// TIA Portal V21 export
// export: Created 2026-11-11T00:48:17.7043043Z, ExportSetting WithDefaults, DisplayName Totally Integrated Automation Portal, DisplayVersion V21 Update 3, DisplayName STEP 7 Professional, DisplayVersion V21 Update 3, DisplayName STEP 7 Safety, DisplayVersion V21, DisplayName Tech WebApplication, DisplayVersion V21, DisplayName WinCC Basic/Comfort/Advanced, DisplayVersion V21 Update 3, DisplayName WinCC Unified, DisplayVersion V21 Update 3
FUNCTION_BLOCK "FB_Scl_sl053"   // FB31, SCL
{ S7_Optimized_Access := 'TRUE' }
VERSION : 0.1
// stored: AutoNumber true, IsIECCheckEnabled false, IsRetainMemResEnabled false, MemoryReserve 100, SetENOAutomatically false, UDAEnableTagReadback false
   VAR_INPUT
      v_req : Bool;
      v_db : DB_ANY;
      v_index : DInt;
   END_VAR
   VAR_OUTPUT
      v_busy : Bool;
      v_done : Bool;
      v_error : Int;
   END_VAR
   VAR_IN_OUT
      v_value : Variant;
   END_VAR
   VAR
      inst { S7_SetPoint := 'True'} : ReadFromArrayDBL;
   END_VAR
BEGIN
   #inst(req := #v_req, db := #v_db, index := #v_index, value := #v_value, busy => #v_busy, done => #v_done, error => #v_error);
END_FUNCTION_BLOCK
